Fanuc KAREL source: KT00946.KL

PROGRAM KT00946
%NOLOCKGROUP
VAR
  ENTRY: INTEGER
  PNAME: STRING[80]
  VNAME: STRING[80]
  STATUS: INTEGER
  VALUE: ARRAY[4] OF REAL
BEGIN
  ENTRY = 0
  PNAME = ''
  VNAME = 'VALUE'
  GET_VAR(ENTRY, PNAME, VNAME, VALUE, STATUS)
END KT00946
